FUNCTION_BLOCK UV_Trojan (* Sistema UV Trojan UV3000Plus (monitoracao Modbus TCP) - HidrycoLib *)
  (* Standard: 61499-2 *)
  (* Version 1.1, 19/10/2026, Hidryco, Hidryco, 1.1: raio do gerador nos canais (REQ_GERADOR com geradorHabilitaCanal1/2 e stsGerador; AnimGeradorCanal1/2 -> STS_CH1/CH2_ANIMACAO_GERADOR). So indicacao: o SCC nao aceita comando. 1.0: Trojan UV3000Plus (SCC M580, servidor Modbus TCP, CP141200010 p.606-611). Campo por symlink ${PATH}: leitura mbR41001..mbR41191 (INT, registro = nome), mbConexao (connStatusInt, 1 = online); escrita mbW40006 (heartbeat bit 1). Somente monitoracao: o SCC nao aceita comandos por rede. *)
  PACKAGE Hidryco.HidrycoLib;
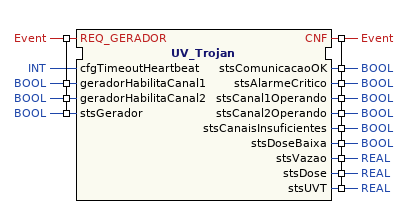
  EVENT_INPUT
    REQ_GERADOR WITH geradorHabilitaCanal1, geradorHabilitaCanal2, stsGerador; (* Planta no gerador e liberacao dos canais (Subestacao) *)
  END_EVENT
  EVENT_OUTPUT
    CNF WITH stsComunicacaoOK, stsAlarmeCritico, stsCanal1Operando, stsCanal2Operando, stsCanaisInsuficientes, stsDoseBaixa, stsVazao, stsDose, stsUVT; (* Status (alarmes na hora, valores a cada 1 s) *)
  END_EVENT
  VAR_INPUT
    cfgTimeoutHeartbeat : INT := 10; (* Tempo sem alternar o heartbeat do SCC para falha de comunicacao (s) *)
    geradorHabilitaCanal1 : BOOL; (* 700-UV-01 (canal 1) liberado para operar com a planta nos geradores *)
    geradorHabilitaCanal2 : BOOL; (* 700-UV-02 (canal 2) liberado para operar com a planta nos geradores *)
    stsGerador : BOOL; (* TRUE = planta alimentada pelos geradores *)
  END_VAR
  VAR_OUTPUT
    stsComunicacaoOK : BOOL; (* Comunicacao Modbus e heartbeat do SCC OK *)
    stsAlarmeCritico : BOOL; (* Alarme comum critico (41001.2) *)
    stsCanal1Operando : BOOL; (* Canal 1 em operacao *)
    stsCanal2Operando : BOOL; (* Canal 2 em operacao *)
    stsCanaisInsuficientes : BOOL; (* Canais saudaveis insuficientes (41003.1) *)
    stsDoseBaixa : BOOL; (* Dose abaixo do alvo (41003.0) *)
    stsVazao : REAL; (* Vazao do sistema no SCC (41005 x fator 41008) *)
    stsDose : REAL; (* Dose equivalente RED (mJ/cm2) *)
    stsUVT : REAL; (* Transmitancia UV (%) *)
  END_VAR
  FBS
    IThis : UV_Trojan_HMI(QI := TRUE);
    plcStart1 : plcStart(Prio := 10);
    Leitura1 : SYMLINKMULTIVARDST_115C998103CD7017B(QI := TRUE, NAME1 := '$${PATH}mbR41001', NAME2 := '$${PATH}mbR41003', NAME3 := '$${PATH}mbR41004', NAME4 := '$${PATH}mbR41005', NAME5 := '$${PATH}mbR41006', NAME6 := '$${PATH}mbR41007', NAME7 := '$${PATH}mbR41008', NAME8 := '$${PATH}mbR41021', NAME9 := '$${PATH}mbR41022', NAME10 := '$${PATH}mbR41031', NAME11 := '$${PATH}mbR41033', NAME12 := '$${PATH}mbR41034', NAME13 := '$${PATH}mbR41035', NAME14 := '$${PATH}mbR41036', NAME15 := '$${PATH}mbR41037'); {SET_ATTRIBUTE(Configuration.GenericFBType.InterfaceParams, Runtime.System#I:=15;VALUE${I$}:INT,INT,INT,INT,INT,INT,INT,INT,INT,INT,INT,INT,INT,INT,INT)}
    Leitura2 : SYMLINKMULTIVARDST_182274139AA51730B(QI := TRUE, NAME1 := '$${PATH}mbR41061', NAME2 := '$${PATH}mbR41062', NAME3 := '$${PATH}mbR41071', NAME4 := '$${PATH}mbR41073', NAME5 := '$${PATH}mbR41074', NAME6 := '$${PATH}mbR41075', NAME7 := '$${PATH}mbR41076', NAME8 := '$${PATH}mbR41077', NAME9 := '$${PATH}mbR41181', NAME10 := '$${PATH}mbR41183', NAME11 := '$${PATH}mbR41185', NAME12 := '$${PATH}mbR41186'); {SET_ATTRIBUTE(Configuration.GenericFBType.InterfaceParams, Runtime.System#I:=12;VALUE${I$}:INT,INT,INT,INT,INT,INT,INT,INT,INT,INT,INT,INT)}
    Leitura3 : SYMLINKMULTIVARDST_15292F208F22048C1(QI := TRUE, NAME1 := '$${PATH}mbR41187', NAME2 := '$${PATH}mbR41189', NAME3 := '$${PATH}mbR41190', NAME4 := '$${PATH}mbR41191'); {SET_ATTRIBUTE(Configuration.GenericFBType.InterfaceParams, Runtime.System#I:=4;VALUE${I$}:INT,INT,INT,INT)}
    Conexao : SYMLINKMULTIVARDST_5A03F112CD5D470(QI := TRUE, NAME1 := '$${PATH}mbConexao'); {SET_ATTRIBUTE(Configuration.GenericFBType.InterfaceParams, Runtime.System#I:=1;VALUE${I$}:INT)}
    Escrita : SYMLINKMULTIVARSRC_5A03F112CD5D470(QI := TRUE, NAME1 := '$${PATH}mbW40006'); {SET_ATTRIBUTE(Configuration.GenericFBType.InterfaceParams, Runtime.System#I:=1;VALUE${I$}:INT)}
    Logica : basicUVTrojan;
    Tick : E_CYCLE(DT := T#1s);
    AlarmeComunicacao : ALARM_BIT(TYPE := 1, ACKTYPE_1 := 2, ACTIVE := TRUE); {SET_ATTRIBUTE(HMI.AlarmText, Sistema UV sem comunicação)} {SET_ATTRIBUTE(HMI.AlarmClass, Warning)}
    AlarmeCritico : ALARM_BIT(TYPE := 1, ACKTYPE_1 := 2, ACTIVE := TRUE); {SET_ATTRIBUTE(HMI.AlarmText, Sistema UV: alarme crítico)}
    AlarmeMaior : ALARM_BIT(TYPE := 1, ACKTYPE_1 := 2, ACTIVE := TRUE); {SET_ATTRIBUTE(HMI.AlarmText, Sistema UV: alarme maior)}
    AlarmeMenor : ALARM_BIT(TYPE := 1, ACKTYPE_1 := 2, ACTIVE := TRUE); {SET_ATTRIBUTE(HMI.AlarmText, Sistema UV: alarme menor)} {SET_ATTRIBUTE(HMI.AlarmClass, Warning)}
    AlarmeLimpeza : ALARM_BIT(TYPE := 1, ACKTYPE_1 := 2, ACTIVE := TRUE); {SET_ATTRIBUTE(HMI.AlarmText, Sistema UV: alarme do sistema de limpeza)} {SET_ATTRIBUTE(HMI.AlarmClass, Warning)}
    AnimGeradorCanal1 : basicCargaGerador(pin_AB02A6BAE011AA16 := TRUE);
    AnimGeradorCanal2 : basicCargaGerador(pin_AB02A6BAE011AA16 := TRUE);
  END_FBS
  EVENT_CONNECTIONS
    plcStart1.FIRST_INIT TO IThis.A0AFE703E8197FF1;
    plcStart1.REDO_INIT TO IThis.A0AFE703E8197FF1;
    IThis.A43DF82B03CDE235 TO Leitura1.INIT;
    Leitura1.INITO TO Leitura2.INIT;
    Leitura2.INITO TO Leitura3.INIT;
    Leitura3.INITO TO Conexao.INIT;
    Conexao.INITO TO Escrita.INIT;
    Escrita.INITO TO Logica.422593B0E0FDF699;
    Logica.E60E8993B78C691A TO Tick.START;
    Logica.E60E8993B78C691A TO AlarmeComunicacao.INIT;
    AlarmeComunicacao.INITO TO AlarmeComunicacao.REQ_INITDATA;
    AlarmeComunicacao.CNF_INITDATA TO AlarmeComunicacao.ACTIVATE;
    AlarmeCritico.INITO TO AlarmeCritico.REQ_INITDATA;
    AlarmeCritico.CNF_INITDATA TO AlarmeCritico.ACTIVATE;
    AlarmeComunicacao.INITO TO AlarmeCritico.INIT;
    AlarmeMaior.INITO TO AlarmeMaior.REQ_INITDATA;
    AlarmeMaior.CNF_INITDATA TO AlarmeMaior.ACTIVATE;
    AlarmeCritico.INITO TO AlarmeMaior.INIT;
    AlarmeMenor.INITO TO AlarmeMenor.REQ_INITDATA;
    AlarmeMenor.CNF_INITDATA TO AlarmeMenor.ACTIVATE;
    AlarmeMaior.INITO TO AlarmeMenor.INIT;
    AlarmeLimpeza.INITO TO AlarmeLimpeza.REQ_INITDATA;
    AlarmeLimpeza.CNF_INITDATA TO AlarmeLimpeza.ACTIVATE;
    AlarmeMenor.INITO TO AlarmeLimpeza.INIT;
    AlarmeLimpeza.INITO TO plcStart1.ACK_FIRST;
    Leitura1.CNF TO Logica.834A2A2E2E7047C9;
    Leitura2.CNF TO Logica.9A75195D93F465A6;
    Leitura3.CNF TO Logica.7AB0ED5945B252F7;
    Conexao.CNF TO Logica.13AC09953D6E2466;
    Tick.EO TO Logica.3A15BE6083DBA891;
    Logica.676B16D752D3B543 TO CNF;
    IThis.3794C9BBA3053F71 TO Logica.E1D341542AF03203;
    Logica.BC8871B735E03A3B TO IThis.EB65E8EFF6E74925;
    Logica.BC8871B735E03A3B TO AlarmeComunicacao.REQ;
    AlarmeComunicacao.IND_1 TO IThis.EB65E8EFF6E74925;
    IThis.3794C9BBA3053F71 TO AlarmeComunicacao.ACK_C1;
    Logica.BC8871B735E03A3B TO AlarmeCritico.REQ;
    AlarmeCritico.IND_1 TO IThis.EB65E8EFF6E74925;
    IThis.3794C9BBA3053F71 TO AlarmeCritico.ACK_C1;
    Logica.BC8871B735E03A3B TO AlarmeMaior.REQ;
    AlarmeMaior.IND_1 TO IThis.EB65E8EFF6E74925;
    IThis.3794C9BBA3053F71 TO AlarmeMaior.ACK_C1;
    Logica.BC8871B735E03A3B TO AlarmeMenor.REQ;
    AlarmeMenor.IND_1 TO IThis.EB65E8EFF6E74925;
    IThis.3794C9BBA3053F71 TO AlarmeMenor.ACK_C1;
    Logica.BC8871B735E03A3B TO AlarmeLimpeza.REQ;
    AlarmeLimpeza.IND_1 TO IThis.EB65E8EFF6E74925;
    IThis.3794C9BBA3053F71 TO AlarmeLimpeza.ACK_C1;
    Logica.581232B93B1DD4EF TO Escrita.REQ;
    REQ_GERADOR TO AnimGeradorCanal1.00789A423C908128;
    REQ_GERADOR TO AnimGeradorCanal2.00789A423C908128;
    Logica.BC8871B735E03A3B TO AnimGeradorCanal1.00789A423C908128;
    Logica.BC8871B735E03A3B TO AnimGeradorCanal2.00789A423C908128;
    AnimGeradorCanal1.D13B80EB42E4132B TO IThis.EB65E8EFF6E74925;
    AnimGeradorCanal2.D13B80EB42E4132B TO IThis.EB65E8EFF6E74925;
  END_CONNECTIONS
  DATA_CONNECTIONS
    Leitura1.VALUE1 TO Logica.2A8FFE90B1F1E261;
    Leitura1.VALUE2 TO Logica.74D7C12CD1DE6A44;
    Leitura1.VALUE3 TO Logica.8842E41C53AAEF18;
    Leitura1.VALUE4 TO Logica.21F26D97BF4440A8;
    Leitura1.VALUE5 TO Logica.72902E44E6AD4B76;
    Leitura1.VALUE6 TO Logica.C4C1A0D0EDACCB0A;
    Leitura1.VALUE7 TO Logica.E6EE9917A3E22159;
    Leitura1.VALUE8 TO Logica.37BB2B157B53007C;
    Leitura1.VALUE9 TO Logica.1D1C7AB0C7D67B87;
    Leitura1.VALUE10 TO Logica.F28C3F14F2F0EC59;
    Leitura1.VALUE11 TO Logica.3C9F79EBC9EDCC30;
    Leitura1.VALUE12 TO Logica.62A97B57D8307687;
    Leitura1.VALUE13 TO Logica.8E79DF9B77C48766;
    Leitura1.VALUE14 TO Logica.A09E5AE1D0AC0328;
    Leitura1.VALUE15 TO Logica.79930D8FEC011FC1;
    Leitura2.VALUE1 TO Logica.DCB5A182CCDF772A;
    Leitura2.VALUE2 TO Logica.12592094A01DFE7B;
    Leitura2.VALUE3 TO Logica.AA0366AAC418F1C1;
    Leitura2.VALUE4 TO Logica.40C89611DD35AFE6;
    Leitura2.VALUE5 TO Logica.45683CE7F872D6EA;
    Leitura2.VALUE6 TO Logica.E7CD76807C7C7229;
    Leitura2.VALUE7 TO Logica.63FBF805A8A252CA;
    Leitura2.VALUE8 TO Logica.FC8DC516B62AEAC6;
    Leitura2.VALUE9 TO Logica.0F7B4990A5DD0A53;
    Leitura2.VALUE10 TO Logica.3C127675843BFB97;
    Leitura2.VALUE11 TO Logica.BADC93940027513E;
    Leitura2.VALUE12 TO Logica.CDE3AED714FCEA41;
    Leitura3.VALUE1 TO Logica.C27D5F866F4B52CE;
    Leitura3.VALUE2 TO Logica.32BC19590FF49687;
    Leitura3.VALUE3 TO Logica.9EC85E4F37DB09DC;
    Leitura3.VALUE4 TO Logica.38575752AD52EF33;
    Conexao.VALUE1 TO Logica.25AA89FA4BD4B0BE;
    cfgTimeoutHeartbeat TO Logica.3DDD936EC9FED321;
    Logica.3F25CD83F3646805 TO stsComunicacaoOK;
    Logica.7B3D3BC0BF1F6804 TO stsAlarmeCritico;
    Logica.018A4B302C939307 TO stsCanal1Operando;
    Logica.6A9501B8C3966D94 TO stsCanal2Operando;
    Logica.DA207E51535047FE TO stsCanaisInsuficientes;
    Logica.309484C904E5427C TO stsDoseBaixa;
    Logica.E7413D0448213082 TO stsVazao;
    Logica.42310D3F28314002 TO stsDose;
    Logica.F778C4FD8D4B5D49 TO stsUVT;
    IThis.DCF094E1991E4C2C TO Logica.ED817AC9D2485697;
    Logica.3F25CD83F3646805 TO IThis.7BF54A23B1B23775;
    Logica.F3F15666596AA2AE TO IThis.2C6EFDE92188C531;
    Logica.C7E90AD487E14A5D TO IThis.FCD86879745E1FE9;
    Logica.C26714600235CB99 TO IThis.C44EE288ADFB5541;
    Logica.8FA1F45CA3D29123 TO IThis.A098053F481CFC62;
    Logica.7B3D3BC0BF1F6804 TO IThis.6D76690FF5D71C8B;
    Logica.DE98D16347DE4799 TO IThis.6D522AE81F4D5A68;
    Logica.8164094A4CD36EEA TO IThis.43B29CCD79780B2F;
    Logica.309484C904E5427C TO IThis.3A1A6E80BF3C33DE;
    Logica.DA207E51535047FE TO IThis.7AADBCAF26F47A9C;
    Logica.E7413D0448213082 TO IThis.FFF98B3E1BCBCADC;
    Logica.42310D3F28314002 TO IThis.FDBA08C3B42F69BA;
    Logica.F778C4FD8D4B5D49 TO IThis.53963A97CABCA69C;
    Logica.5340B3252E0ED0C2 TO IThis.56104A8898640B3F;
    Logica.E38B6D26792FBA9C TO IThis.A82556935290A563;
    Logica.ED012D70C0C16781 TO IThis.478DB10CB39141B5;
    Logica.20066233F2045EE6 TO IThis.57CB5ADF0C170B7B;
    Logica.018A4B302C939307 TO IThis.F83E7A2124F4CD00;
    Logica.7A0641EEBAA0BD94 TO IThis.B78368F8D4B5B8BF;
    Logica.0D626260960EF09F TO IThis.27D9BF65E041688B;
    Logica.7D933C7D3B13940F TO IThis.C6DFB64F5EEF40B2;
    Logica.4CD3F240D079AA40 TO IThis.801CE9A9AAA0241E;
    Logica.0CE6BC70DC8F15BE TO IThis.E33BE408E47EE7AE;
    Logica.174494CCD7E64F21 TO IThis.1800066AD3EE1A6F;
    Logica.67075D43B5C92663 TO IThis.E1925219F6A86BD5;
    Logica.273C0A990E1C720E TO IThis.53A2F2B1D4625D7E;
    Logica.77DD43FE18278936 TO IThis.5DFCCDCD258F4DA7;
    Logica.27271CF9D3195869 TO IThis.7B87E3644EEB05B2;
    Logica.B10278E129C430C7 TO IThis.7F726B1E9B28435A;
    Logica.FB18D177E4913472 TO IThis.90607E9D75E08886;
    Logica.6A9501B8C3966D94 TO IThis.4B2546588D516929;
    Logica.0BD8C968EFFF6E26 TO IThis.219E940EBB37CB9F;
    Logica.FDE4D5ABB944D921 TO IThis.66D20250FAF8B0D2;
    Logica.C689C70844359B1B TO IThis.0D4CD33E7A5FED20;
    Logica.A862306AB43ACCAC TO IThis.D797CA5E010B507E;
    Logica.486502E514D94D6E TO IThis.AC2B42B37D274536;
    Logica.B89234385FB47CE2 TO IThis.EFE2B134242D36EE;
    Logica.F839FAAF949206F4 TO IThis.DAA220F8CC7F1283;
    Logica.7DCC6373C5D04F35 TO IThis.645E0F0EE2E39F37;
    Logica.AD3A738821D8DF93 TO IThis.DB675BBD907AC9EE;
    Logica.F789DC280B22B5EE TO IThis.0412DE6AC3839F8E;
    Logica.4A326CAA691F5553 TO IThis.28A2DEA0B8A3C68F;
    Logica.6D744FDCA439A4CB TO IThis.4C09D7B13FFF9CC0;
    Logica.D651FFE2071B98FA TO IThis.B4B1F56FDD35CCD6;
    Logica.2E6C286340FF1EC6 TO IThis.39080BE048FC6C3D;
    Logica.7E399129E7E35FF1 TO IThis.CE3E682CAF26D787;
    Logica.5CFCA8DB00DAD867 TO IThis.042BD5540060F137;
    Logica.521A383470437976 TO IThis.CD66B2349BEA8385;
    Logica.AFCBCA6415E3903D TO IThis.F553003F93B6F662;
    Logica.747FEBC2833DFCB0 TO IThis.B8B36C9FEDA67431;
    Logica.C7E90AD487E14A5D TO AlarmeComunicacao.INP;
    AlarmeComunicacao.STATE_1 TO IThis.C798321CD45B4534;
    Logica.7B3D3BC0BF1F6804 TO AlarmeCritico.INP;
    AlarmeCritico.STATE_1 TO IThis.DEF003E8B8A46241;
    Logica.8FA1F45CA3D29123 TO AlarmeMaior.INP;
    AlarmeMaior.STATE_1 TO IThis.DB2738DEE3749551;
    Logica.C26714600235CB99 TO AlarmeMenor.INP;
    AlarmeMenor.STATE_1 TO IThis.22DB8D49A045D74A;
    Logica.DE98D16347DE4799 TO AlarmeLimpeza.INP;
    AlarmeLimpeza.STATE_1 TO IThis.9DC737B08AFBDB3E;
    Logica.06946B36B49CCADC TO Escrita.VALUE1;
    geradorHabilitaCanal1 TO AnimGeradorCanal1.E98CC3FC79967C8B;
    geradorHabilitaCanal2 TO AnimGeradorCanal2.E98CC3FC79967C8B;
    stsGerador TO AnimGeradorCanal1.9DDD74C1F0C45B78;
    stsGerador TO AnimGeradorCanal2.9DDD74C1F0C45B78;
    Logica.018A4B302C939307 TO AnimGeradorCanal1.92CF573A93E227B1;
    Logica.6A9501B8C3966D94 TO AnimGeradorCanal2.92CF573A93E227B1;
    AnimGeradorCanal1.87DFF1D389B6D369 TO IThis.6328E94C56C87F6C;
    AnimGeradorCanal2.87DFF1D389B6D369 TO IThis.6F057DB5A9F534BA;
  END_CONNECTIONS
END_FUNCTION_BLOCK
